FUNCTION_BLOCK "Tgp_ComponentEffect"
{ S7_Optimized_Access := 'TRUE' }
VERSION : 0.1
VAR_INPUT
 Enable : Bool;
END_VAR
VAR_OUTPUT
 Active : Bool;
END_VAR
VAR
 RetainedMarker : Int := 17;
END_VAR
BEGIN
 #Active := #Enable;
END_FUNCTION_BLOCK

DATA_BLOCK "Tgp_ComponentEffect_DB"
{ S7_Optimized_Access := 'TRUE' }
VERSION : 0.1
"Tgp_ComponentEffect"
BEGIN
 RetainedMarker := 42;
END_DATA_BLOCK
